Staubli VAL3: loadingPage.pgx

public program loadingPage()
begin
  userPage("loading")
  delay(0)
end
